// TwinCAT 3 PLC project VISU_plc
// ProgramVersion: 3.1.4026.25
// libraries:
//   Tc2_Standard, * (Beckhoff Automation GmbH)
//   Tc2_System, * (Beckhoff Automation GmbH)
//   Tc3_Module, * (Beckhoff Automation GmbH)
// project tree:
//   DUTs/ E_Ingredient_type.TcDUT, E_Prod_Status.TcDUT, E_Prod_Type.TcDUT, ST_PLC_To_VisuPLC.TcDUT, ST_Prod_Ingredient.TcDUT, ST_VisuPLC_To_PLC.TcDUT
//   / GlobalTextList.TcGTLO, PlcTask.TcTTO, VisualizationManager.TcVMO (not stored), VISU_TASK.TcTTO
//   GVLs/ g_HMI_Panel.TcGVL
//   POUs/ MAIN.TcPOU
//   VISUs/ vis_Dissolve.TcVIS, vis_ProgressBar.TcVIS
// (motion and I/O tree: see PLC project plc)
// real-time tasks:
//   TASK PlcTask: cycle T#10ms, priority 20, ADS port 350
//   TASK PlcTask_Recipe: cycle T#300ms, priority 14, ADS port 351
//   TASK PlcTask1: cycle T#10ms, priority 21, ADS port 352
//   TASK VISU_TASK: cycle T#200000us, priority 30, ADS port 353
// variable links:

CONFIGURATION VISU_plc
    RESOURCE PLC ON TwinCAT3
        TASK PlcTask(INTERVAL := T#10ms, PRIORITY := 21);
        TASK VISU_TASK(INTERVAL := T#200000us, PRIORITY := 30);
        PROGRAM MAIN WITH PlcTask : MAIN;
        PROGRAM VisuElems_Visu_Prg WITH VISU_TASK : VisuElems.Visu_Prg;
    END_RESOURCE
END_CONFIGURATION

// ---- DUTs/E_Ingredient_type.TcDUT
{attribute 'qualified_only'}
{attribute 'strict'}
TYPE E_Ingredient_type :
(
	eNone := 0,
	eWater,
	ePowder,
	eOil
);
END_TYPE

// ---- DUTs/E_Prod_Status.TcDUT
{attribute 'qualified_only'}
{attribute 'strict'}
TYPE E_Prod_Status :
(
	Not_Active := 0,
	Activation_Pending,
	Activation_Pending_Shift, // to shift UTC 
	Active
);
END_TYPE

// ---- DUTs/E_Prod_Type.TcDUT
{attribute 'qualified_only'}
{attribute 'strict'}
TYPE E_Prod_Type :
(
	Marinade := 0,
	Color
);
END_TYPE

// ---- DUTs/ST_PLC_To_VisuPLC.TcDUT
TYPE ST_PLC_To_VisuPLC :
STRUCT
	lifeBit: BOOL;
	
// General
	Description				: STRING(30);
	prodType				: E_Prod_Type;	
	RPM_FeedBack			: REAL;
	Flow_FeedBack			: REAL;
	fBlendingPercenatge		: DINT;
	
// Component
	arr_Component			: ARRAY [1..10] OF ST_Prod_Ingredient;

	iActual_Component		: INT;
	bDissolving_Active		: BOOL;
	bBlending_Active		: BOOL;
	bMainPause_Active		: BOOL;

END_STRUCT
END_TYPE

// ---- DUTs/ST_Prod_Ingredient.TcDUT
TYPE ST_Prod_Ingredient :
STRUCT
	sDescription		: STRING:= 'Ingredient Name';
	eIngredientType		: E_Ingredient_type;
	rWeight				: REAL; // kg
	rWeightPercentage	: REAL;
	rFlowRate_Dissolving: REAL;
	rFlowRate_Blending	: REAL;
	tBlendingDuration	: TIME;

END_STRUCT
END_TYPE

// ---- DUTs/ST_VisuPLC_To_PLC.TcDUT
TYPE ST_VisuPLC_To_PLC :
STRUCT
	lifeBit: BOOL;
	
	RPM_setPoint: REAL;
	
	bPauseTriBlender: BOOL;
	
	bActualComponentDisolving_Done: BOOL;



END_STRUCT
END_TYPE

// ---- GVLs/g_HMI_Panel.TcGVL
//{attribute 'qualified_only'}
VAR_GLOBAL
	stVisuPLC_To_PLC		AT %MB1000 : ST_VisuPLC_To_PLC;
	stPLC_To_VisuPLC		AT %MB2000 : ST_PLC_To_VisuPLC;
	
	q_stVisuPLC_To_PLC		AT %Q* : ST_VisuPLC_To_PLC;
	i_stPLC_To_VisuPLC		AT %I* : ST_PLC_To_VisuPLC;
END_VAR

// ---- POUs/MAIN.TcPOU
PROGRAM MAIN
VAR
	k: REAL;
	ton_Life: TON;
	memo_last_component_Index: INT;
	ton_BlendingTime: TON;
	tBlendingRemainTime: DINT;
	fBlendingPercenatge: DINT;
	ptTemp: DINT;
	realTemp: REAL;
	iProgressBarOfset: DINT;
	iActualComponentDisolving_Done_lifetime: INT;
	ftDissolvingActive: F_TRIG;
END_VAR

k:=k+1;

//g_HMI_Panel.stVisuPLC_To_PLC.RPM_setPoint:=k;

ton_Life(PT:=T#1S, IN:=NOT ton_Life.Q);
IF ton_Life.ET>T#0.5S THEN;
	g_HMI_Panel.stVisuPLC_To_PLC.lifeBit:=TRUE;
ELSE;
	g_HMI_Panel.stVisuPLC_To_PLC.lifeBit:=FALSE;
END_IF


IF memo_last_component_Index <> stPLC_To_VisuPLC.iActual_Component THEN;
	IF stPLC_To_VisuPLC.iActual_Component>=1 AND stPLC_To_VisuPLC.iActual_Component<=10 THEN;
		stVisuPLC_To_PLC.RPM_setPoint:=stPLC_To_VisuPLC.arr_Component[stPLC_To_VisuPLC.iActual_Component].rFlowRate_Dissolving;
		ton_BlendingTime(PT:=g_HMI_Panel.stPLC_To_VisuPLC.arr_Component[stPLC_To_VisuPLC.iActual_Component].tBlendingDuration);
	ELSE;
		stVisuPLC_To_PLC.RPM_setPoint:=0;
	END_IF	
	memo_last_component_Index:= stPLC_To_VisuPLC.iActual_Component;
	g_HMI_Panel.stVisuPLC_To_PLC.bActualComponentDisolving_Done:=FALSE;
END_IF


ton_BlendingTime();
IF g_HMI_Panel.stPLC_To_VisuPLC.bBlending_Active THEN;
	ton_BlendingTime.IN:=TRUE;
	tBlendingRemainTime:=TIME_TO_DINT(ton_BlendingTime.PT - ton_BlendingTime.ET);
ELSE;
	ton_BlendingTime.IN:=FALSE;
END_IF

ptTemp:=TIME_TO_DINT(ton_BlendingTime.PT);
IF ton_BlendingTime.PT<>T#0S THEN;
	realTemp:=(DINT_TO_REAL(tBlendingRemainTime)/DINT_TO_REAL(ptTemp)*100.0);
	fBlendingPercenatge:=TRUNC(realTemp);
END_IF

iProgressBarOfset:=TRUNC(stPLC_To_VisuPLC.iActual_Component*37.2);

ftDissolvingActive(CLK:=g_HMI_Panel.stPLC_To_VisuPLC.bDissolving_Active);
IF ftDissolvingActive.Q THEN;
	g_HMI_Panel.stVisuPLC_To_PLC.bActualComponentDisolving_Done:=FALSE;
END_IF

(*
IF iActualComponentDisolving_Done_lifetime>0 THEN;
	iActualComponentDisolving_Done_lifetime:=0;
	g_HMI_Panel.stVisuPLC_To_PLC.bActualComponentDisolving_Done:=FALSE;
END_IF
IF g_HMI_Panel.stVisuPLC_To_PLC.bActualComponentDisolving_Done THEN;
	iActualComponentDisolving_Done_lifetime:=iActualComponentDisolving_Done_lifetime+1;	
END_IF
*)

END_PROGRAM

// ---- GlobalTextList.TcGTLO
TEXTLIST GlobalTextList
  443 = '\tRecipe name: %s'
  556 = '  %4.0f rpm'
  322 = '  %4.1f liter/h'
  448 = '  %4.1f liter/hour'
  487 = '  %4.1f rpm'
  971 = ' Recipe type: %s'
  989 = '%'
  341 = '%4.0f'
  937 = '%4.0f rpm'
  470 = '%4.1f'
  826 = '%4.2f'
  187 = '%4f'
  36 = '%4f rpm'
  155 = '%d'
  720 = '%d rpm'
  479 = '%f4.1'
  964 = 'Component Description'
  391 = 'DONE'
  42 = 'DOWN'
  703 = 'Flow Rate'
  584 = 'Flow [RPM]'
  988 = 'main Pause active'
  485 = 'Pause'
  476 = 'Play'
  668 = 'Recipe name: %s'
  33 = 'Type'
  515 = 'UP'
  417 = 'Weight'
  758 = 'Weight Percentage'
  631 = 'Weight [kg]'
END_TEXTLIST

// ---- VISUs/vis_Dissolve.TcVIS
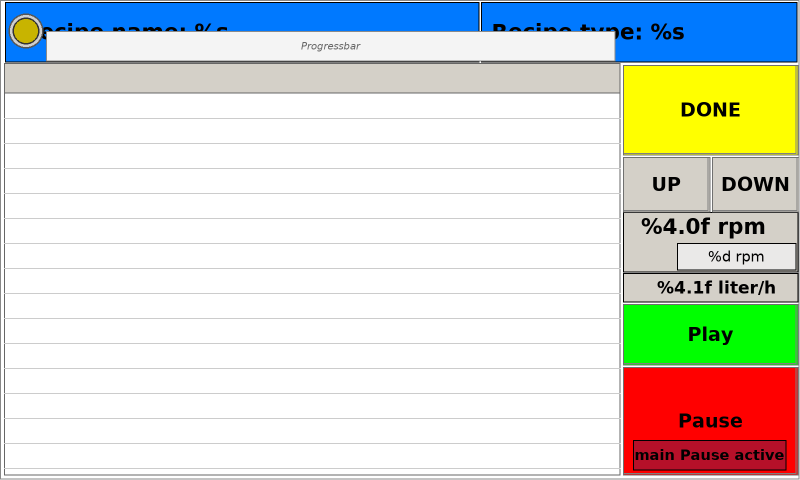
VISUALIZATION vis_Dissolve  // 800x480
VAR_IN_OUT
	
END_VAR

VAR
	lacal_bool: BOOL:=TRUE;
END_VAR
    Table (4,63 616x412), data array: stPLC_To_VisuPLC.arr_Component
        p3854506369: stPLC_To_VisuPLC.arr_Component[INDEX].sDescription
        p1892666644: stPLC_To_VisuPLC.arr_Component[INDEX].eIngredientType
        p338671338: stPLC_To_VisuPLC.arr_Component[INDEX].rWeight
        p2170511999: stPLC_To_VisuPLC.arr_Component[INDEX].rWeightPercentage
        p3723444502: stPLC_To_VisuPLC.arr_Component[INDEX].rFlowRate_Dissolving
        p1218418051: stPLC_To_VisuPLC.arr_Component[INDEX].rFlowRate_Blending
        p746581629: stPLC_To_VisuPLC.arr_Component[INDEX].tBlendingDuration
        p2232123230: Component Description
        p1755163831: Weight [kg]
        p4092479075: %
        p2237128397: Flow [RPM]
        p1137915858: stPLC_To_VisuPLC.iActual_Component
    Rectangle (623,212 175x60), "%4.0f rpm", text variable: g_HMI_Panel.stVisuPLC_To_PLC.RPM_setPoint
    Button (623,157 87x55), "UP", input disabled if: NOT g_HMI_Panel.stPLC_To_VisuPLC.bDissolving_Active
        OnMouseDown: execute {
            g_HMI_Panel.stVisuPLC_To_PLC.RPM_setPoint:=
            g_HMI_Panel.stVisuPLC_To_PLC.RPM_setPoint+50;
            IF g_HMI_Panel.stVisuPLC_To_PLC.RPM_setPoint>2500 THEN;
            	g_HMI_Panel.stVisuPLC_To_PLC.RPM_setPoint:=2500;
            END_IF
        }
    Button (712,157 87x55), "DOWN", input disabled if: NOT g_HMI_Panel.stPLC_To_VisuPLC.bDissolving_Active
        OnMouseDown: execute {
            g_HMI_Panel.stVisuPLC_To_PLC.RPM_setPoint:=
            g_HMI_Panel.stVisuPLC_To_PLC.RPM_setPoint-50;
            IF g_HMI_Panel.stVisuPLC_To_PLC.RPM_setPoint<300 THEN;
            	g_HMI_Panel.stVisuPLC_To_PLC.RPM_setPoint:=300;
            END_IF
        }
    Rectangle (5,2 474x60), "Recipe name: %s", text variable: g_HMI_Panel.stPLC_To_VisuPLC.Description
    Lamp1 (6,11 40x40), variable: g_HMI_Panel.stPLC_To_VisuPLC.lifeBit, style: Lamp-Lamp1-Yellow
    Rectangle (677,243 119x27), "%d rpm", text variable: g_HMI_Panel.stPLC_To_VisuPLC.RPM_FeedBack
    Rectangle (481,2 316x60), "Recipe type: %s", text variable: g_HMI_Panel.stPLC_To_VisuPLC.prodType
    Button (623,367 175x108), "Pause", colour toggle: g_HMI_Panel.stVisuPLC_To_PLC.bPauseTriBlender, pressed state: g_HMI_Panel.stVisuPLC_To_PLC.bPauseTriBlender, input disabled if: g_HMI_Panel.stVisuPLC_To_PLC.bPauseTriBlender OR NOT g_HMI_Panel.stPLC_To_VisuPLC.bDissolving_Active
        toggle g_HMI_Panel.stVisuPLC_To_PLC.bPauseTriBlender
    Button (623,304 175x61), "Play", colour toggle: NOT g_HMI_Panel.stVisuPLC_To_PLC.bPauseTriBlender, pressed state: NOT g_HMI_Panel.stVisuPLC_To_PLC.bPauseTriBlender, input disabled if: NOT g_HMI_Panel.stVisuPLC_To_PLC.bPauseTriBlender
        toggle g_HMI_Panel.stVisuPLC_To_PLC.bPauseTriBlender
    Button (623,65 175x90), "DONE", input disabled if: NOT g_HMI_Panel.stPLC_To_VisuPLC.bDissolving_Active OR g_HMI_Panel.stVisuPLC_To_PLC.bPauseTriBlender
        OnMouseClick: execute { g_HMI_Panel.stVisuPLC_To_PLC.bActualComponentDisolving_Done:=TRUE; }
    Rectangle (3,100 618x378)
    Frame (46,31 569x30), invisible if: NOT g_HMI_Panel.stPLC_To_VisuPLC.bBlending_Active
        shows vis_ProgressBar()
        p2738717112: MAIN.iProgressBarOfset
    Rectangle (623,273 175x29), "%4.1f liter/h", text variable: g_HMI_Panel.stPLC_To_VisuPLC.Flow_FeedBack
    Rectangle (633,440 153x30), "main Pause active", invisible if: NOT g_HMI_Panel.stPLC_To_VisuPLC.bMainPause_Active
END_VISUALIZATION

// ---- VISUs/vis_ProgressBar.TcVIS
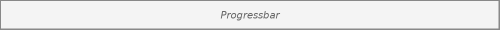
VISUALIZATION vis_ProgressBar  // 500x30
    Progressbar (0,0 500x30), variable: g_HMI_Panel.stPLC_To_VisuPLC.fBlendingPercenatge
END_VISUALIZATION
